Fanuc KAREL source: KO00121.KL

PROGRAM KO00121
%NOLOCKGROUP
VAR
  A: ARRAY[2] OF SHORT
  B: INTEGER
  OUT: INTEGER
BEGIN
  A[1] = 1
  B = 2
  OUT = ATAN2(A[1], B)
END KO00121
